ADAPTER CONVEYOR_HS (* Adapter Interface *)
  (* Standard: 61499-1 *)
  (* Version 0.0, 7/2/2026 *)
  PACKAGE Main;
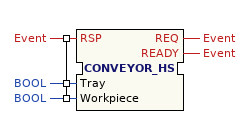
  EVENT_INPUT
    RSP WITH Workpiece, Tray; (* Response from Socket *)
  END_EVENT
  EVENT_OUTPUT
    REQ; (* Confirmation from Plug *)
    READY; (* Indication from Plug *)
  END_EVENT
  VAR_INPUT
    Tray : BOOL; (* Request Data from Socket *)
    Workpiece : BOOL; (* Response Data from Socket *)
  END_VAR
  SERVICE SOCKET/PLUG
    SEQUENCE request_confirm
      SOCKET.REQ(Tray) -> PLUG.REQ(Tray);
      PLUG.REQ(CNFD) -> SOCKET.REQ(CNFD);
    END_SEQUENCE
    SEQUENCE indication_response
      PLUG.READY(INDD) -> SOCKET.READY(INDD);
      SOCKET.RSP(Workpiece) -> PLUG.RSP(Workpiece);
    END_SEQUENCE
  END_SERVICE
END_ADAPTER
